(* PLC project Robin example project, CODESYS CODESYS V3.5 SP15, author pdcribeiro *)
(* stored: creationDateTime 2020-03-17T12:31:34.2855802, version 0.0.1, modificationDateTime 2020-03-17T12:31:34.2481636, organization INESC TEC *)
(* An example project for the Robin library.

https://github.com/ScalABLE40/robin *)

TYPE TestStruct : STRUCT
  var_bool : BOOL;
  var_byte : BYTE;
  var_int16 : INT;
  var_uint64 : ULINT;
  var_float32 : REAL;
  var_float64 : LREAL;
  var_string : STRING;
  var_pose : Pose;
  var_struct_array : ARRAY[1..2] OF ByteMultiArray;
  {attribute 'robin_var_len'}
  var_struct_varlen_array : ARRAY[1..2] OF ByteMultiArray;
END_STRUCT;
END_TYPE

PROGRAM ROS_PRG
  VAR_INPUT
    bool_to_ros : BOOL;
    double_to_ros : LREAL;
    string_to_ros : STRING;
    {attribute 'robin_var_len'}
    string_varlen_array_to_ros : ARRAY[1..5] OF STRING;
    struct1_to_ros : TestStruct;
    struct2_array_to_ros : ARRAY[1..2] OF AccelStamped;
    rosmsg_to_ros : AccelStamped;
  END_VAR
  VAR_OUTPUT
    bool_to_codesys : BOOL;
    double_to_codesys : LREAL;
    string_to_codesys : STRING;
    {attribute 'robin_var_len'}
    string_varlen_array_to_codesys : ARRAY[1..5] OF STRING;
    struct1_to_codesys : TestStruct;
    struct2_array_to_codesys : ARRAY[1..2] OF AccelStamped;
    rosmsg_to_codesys : AccelStamped;
  END_VAR
  VAR
    robin : Robin;
  END_VAR

                    // instancing Robin class
robin();

//////////////////////////////////////////////////////////////////////////////////////////////////////////////////////////////////////////
//																																		//
//												READ - robin.read(<topic_name>, <variable>)												//
//																																		//
//////////////////////////////////////////////////////////////////////////////////////////////////////////////////////////////////////////
// DEBUG: rostopic pub /bool_to_codesys std_msgs/Bool "data: true/false"
robin.read('bool_to_codesys', bool_to_codesys);

// DEBUG: rostopic pub /double_to_codesys std_msgs/Float64 "data: 42.0"
robin.read('double_to_codesys', double_to_codesys);

// DEBUG: rostopic pub /string_to_codesys std_msgs/String "data: 'hello world!'"
robin.read('string_to_codesys', string_to_codesys);

// DEBUG: rostopic pub /string_varlen_array_to_codesys robin_bridge/StringVarLenArray "{data:[str1, str2, str3, str4, str5]}"
robin.read('string_varlen_array_to_codesys', string_varlen_array_to_codesys);

// DEBUG: rostopic pub /struct1_to_codesys robin_bridge/TestStruct "var_bool: false var_byte: 0 <...>"
robin.read('struct1_to_codesys', struct1_to_codesys);

// DEBUG: rostopic pub /struct2_array_to_codesys robin_bridge/AccelStampedArray "data: - header: <...> -header: <...>"
robin.read('struct2_array_to_codesys', struct2_array_to_codesys);

// DEBUG: rostopic pub /rosmsg_to_ros robin_bridge/AccelStamped "data: - header: <...> -header: <...>"
robin.read('rosmsg_to_codesys', rosmsg_to_codesys);


//////////////////////////////////////////////////////////////////////////////////////////////////////////////////////////////////////////
//																																		//
//												WRITE - robin.write(<topic_name>, <variable>)											//
//																																		//
//////////////////////////////////////////////////////////////////////////////////////////////////////////////////////////////////////////

robin.write('bool_to_ros', bool_to_ros);
robin.write('double_to_ros', double_to_ros);
robin.write('string_to_ros', string_to_ros);
robin.write('string_varlen_array_to_ros', string_varlen_array_to_ros);
robin.write('struct1_to_ros', struct1_to_ros);
robin.write('struct2_array_to_ros', struct2_array_to_ros);
robin.write('rosmsg_to_ros', rosmsg_to_ros);


                  
END_PROGRAM

PROGRAM MAIN

                    (*ROS_PRG.double_to_ros := ROS_PRG.double_to_codesys;
ROS_PRG.string_varlen_array_to_ros := ROS_PRG.string_varlen_array_to_codesys;
ROS_PRG.struct1_to_ros := ROS_PRG.struct1_to_codesys;
ROS_PRG.struct2_array_to_ros := ROS_PRG.struct2_array_to_codesys;*)

                  
END_PROGRAM

CONFIGURATION Device
  RESOURCE Application ON PLC
    TASK MainTask(INTERVAL := T#10ms, PRIORITY := 1);
    PROGRAM MAIN WITH MainTask : MAIN;
    PROGRAM ROS_PRG WITH MainTask : ROS_PRG;
  END_RESOURCE
END_CONFIGURATION

CONFIGURATION SoftMotion General Axis Pool
END_CONFIGURATION
